FUNCTION_BLOCK ValidateType
  (* Standard: 61499-1; Description: Copyright (c) 2026 Martin Erich Jobst This program and the accompanying materials are made available under the terms of the Eclipse Public License 2.0 which is available at https://www.eclipse.org/legal/epl-2.0/ SPDX-License-Identifier: EPL-2.0 *)
  (* Version 1.0, 2026-11-18, Martin Jobst *)
  PACKAGE lib::TypedConfigureableObject;
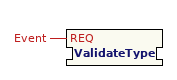
  EVENT_INPUT
    REQ;
  END_EVENT
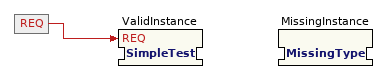
  FBS
    ValidInstance : lib::TypedConfigureableObject::support::SimpleTest;
    MissingInstance : MissingType;
  END_FBS
  EVENT_CONNECTIONS
    REQ TO ValidInstance.REQ;
  END_CONNECTIONS
END_FUNCTION_BLOCK
